screen "Settings" 480x272, template "Template_1"
   TextField "Text_1" at 6,2 size 300x22; Text 'LCP-01 Settings'
   TextField "Text_2" at 330,3 size 146x20; Text 'E-STOP / RESET'
      Visibility <- "Sys_Alm_EStop"
   Button "Button_1" at 2,236 size 76x34; TextOff 'Overview'
      on Press: ActivateScreen("Root screen", 0)
   Button "Button_2" at 82,236 size 76x34; TextOff 'BR01'
      on Press: ActivateScreen("BR01", 0)
   Button "Button_3" at 162,236 size 76x34; TextOff 'BR02'
      on Press: ActivateScreen("BR02", 0)
   Button "Button_4" at 242,236 size 76x34; TextOff 'Scrubber'
      on Press: ActivateScreen("Scrubber", 0)
   Button "Button_5" at 322,236 size 76x34; TextOff 'Alarms'
      on Press: ActivateScreen("Alarms", 0)
   Button "Button_6" at 402,236 size 76x34; TextOff 'Settings'
      on Press: ActivateScreen("Settings", 0)
   TextField "Text_3" at 8,30 size 110x18; Text 'Setting'
   TextField "Text_4" at 120,30 size 76x18; Text 'New'
   TextField "Text_5" at 200,30 size 90x18; Text 'Range'
   TextField "Text_6" at 292,30 size 76x18; Text 'Accepted'
   TextField "Text_7" at 8,50 size 112x20; Text 'Stop at C'
   IOField "IOField_1" at 120,50 size 76x20; FormatPattern s99999
      ProcessValue <- "Par_SP"
   TextField "Text_8" at 200,50 size 90x20; Text '40.0 - 90.0'
   IOField "IOField_2" at 292,50 size 76x20; FormatPattern s99999
      ProcessValue <- "Par_SP_V"
   TextField "Text_9" at 8,72 size 112x20; Text 'Restart below C'
   IOField "IOField_3" at 120,72 size 76x20; FormatPattern s99999
      ProcessValue <- "Par_HYST"
   TextField "Text_10" at 200,72 size 90x20; Text '3.0 - 10.0'
   IOField "IOField_4" at 292,72 size 76x20; FormatPattern s99999
      ProcessValue <- "Par_HYST_V"
   TextField "Text_11" at 8,94 size 112x20; Text '2nd stage below C'
   IOField "IOField_5" at 120,94 size 76x20; FormatPattern s99999
      ProcessValue <- "Par_STG"
   TextField "Text_12" at 200,94 size 90x20; Text '5.0 - 30.0'
   IOField "IOField_6" at 292,94 size 76x20; FormatPattern s99999
      ProcessValue <- "Par_STG_V"
   TextField "Text_13" at 8,116 size 112x20; Text 'Start time ms'
   IOField "IOField_7" at 120,116 size 76x20; FormatPattern s9999999
      ProcessValue <- "Par_TStart"
   TextField "Text_14" at 200,116 size 90x20; Text '90000 - 300000'
   IOField "IOField_8" at 292,116 size 76x20; FormatPattern s9999999
      ProcessValue <- "Par_TStart_V"
   TextField "Text_15" at 8,138 size 112x20; Text 'Drain open ms'
   IOField "IOField_9" at 120,138 size 76x20; FormatPattern s9999999
      ProcessValue <- "Par_TDrnOn"
   TextField "Text_16" at 200,138 size 90x20; Text '1000 - 30000'
   IOField "IOField_10" at 292,138 size 76x20; FormatPattern s9999999
      ProcessValue <- "Par_TDrnOn_V"
   TextField "Text_17" at 8,160 size 112x20; Text 'Drain close ms'
   IOField "IOField_11" at 120,160 size 76x20; FormatPattern s9999999
      ProcessValue <- "Par_TDrnOff"
   TextField "Text_18" at 200,160 size 90x20; Text '0 - 60000'
   IOField "IOField_12" at 292,160 size 76x20; FormatPattern s9999999
      ProcessValue <- "Par_TDrnOff_V"
   TextField "Text_19" at 8,182 size 112x20; Text 'Drain max ms'
   IOField "IOField_13" at 120,182 size 76x20; FormatPattern s9999999
      ProcessValue <- "Par_TDrnMax"
   TextField "Text_20" at 200,182 size 90x20; Text '60000 - 3600000'
   IOField "IOField_14" at 292,182 size 76x20; FormatPattern s9999999
      ProcessValue <- "Par_TDrnMax_V"
   TextField "Text_21" at 372,52 size 104x54; Text 'Raising heat applies after STOP + START.'
   Circle "Circle_1" at 372,117 size 12x12
      Appearance <- "BR01_ParPending"
   TextField "Text_22" at 388,114 size 88x18; Text 'BR01 pending'
   Circle "Circle_2" at 372,137 size 12x12
      Appearance <- "BR02_ParPending"
   TextField "Text_23" at 388,134 size 88x18; Text 'BR02 pending'
   TextField "Text_24" at 8,208 size 360x20; Text 'Setting rejected: out of range (RESET to clear)'
      Visibility <- "Sys_Alm_ParRejected"
   TextField "Text_25" at 372,160 size 104x40; Text 'Settings need log-on (user Engineer).'
*)